(* Logix 5000 project; controller R400_500_XLS vendor 1 type 14 code 216 rev 31.11; software revision 31.01; part 14 of 32 *)
(* tags used below, declared in another part *)
   Abort1 : DINT;   // Not Used
   Alarm : SINT;   // Wait 3 seconds
   AlarmAcked : BOOL;   // Alarm has been acked
   bAlrm : BOOL[64];
   bChangeFromNonHeatedToHeated : BOOL;
   Chem_Pump : UDT_CHEM_PUMP[4];   // Chemical Pump flow rate
   CURRENT_CYCLE : DINT;
   CycExcBuffer : UDT_CYCLE;
   CycleModifBuffer : UDT_CYCLE;
   Cycles : UDT_CYCLE[11];
   DESCALER : SINT;
   ENVIRO_CARE : SINT;
   EXTRA_CARE : SINT;
   FC83_AutoSpeed : BOOL;   // Cycle pump speed selection
   FC83_AutoWtrLevel : BOOL;   // Cycle water level selection
   FC83_CyclePerm : BOOL;   // Cycle permission selection
   FC83_ONS : SINT;
   Inj_Cond : SINT;   // Conductivity injection based steps
   Inj_Time : SINT;   // Time based chemical injection steps
   M : DINT[5];   // Memory Bits
   Neutral : SINT;
   NeutralizantPump : SINT;
   NeutralizationInjTime : DINT;
   NeutralizationPhaseRequired : BOOL;
   NeutralizationRecircTime : DINT;
   ONS_WSH35 : SINT;
   PLASTIC_CARE : SINT;
   PreWash_Select : BOOL;
   PrewashIndex : SINT;   // Index of the selected pre-wash treatment
   RINSE_CARE : SINT;
   RinseIndex : SINT;
   Run : DINT;
   STANDARD : SINT;
   String : STRING[50];   // String
   Supervisor : DINT;
   Tmr : TIMER[107];
   Trt_Wsh : DINT;
   USER_DEFINED_10 : SINT;
   USER_DEFINED_11 : SINT;
   USER_DEFINED_7 : SINT;
   USER_DEFINED_8 : SINT;
   USER_DEFINED_9 : SINT;
   VolumeInjected_ML : REAL;
   VolumeNeutralizer : REAL;
   WashIndex : SINT;
   WshExcBuffer : UDT_WASH;
   cfgPrewashWport : SINT;
   CycleName : STRING[12];
   CyclePtr : DINT;   // Cycle Pointeur
   I_Chm_1_Lvl_Sw : BOOL;   // Chemical Pump #1 level switch
   I_Chm_2_Lvl_Sw : BOOL;   // Chemical Pump #2 level switch
   I_Chm_3_Lvl_Sw : BOOL;   // Chemical Pump #3 level switch
   I_Chm_4_Lvl_Sw : BOOL;   // Chemical Pump #4 level switch
   NumInputReal : UDT_NUMERIC_INPUT_REAL[17];
   Screen_Ctrl : DINT;   // PLC Screen Request
   SelChemNeutralizer : UDT_SELECTOR[5];
   Selector : UDT_SELECTOR[25];   // Piloted list selector
   Tpb : DINT[11];
   TpbImage : DINT[11];
   Unit : Hrdwre;   // Unit Configuration
(* MainProgram, continued *)

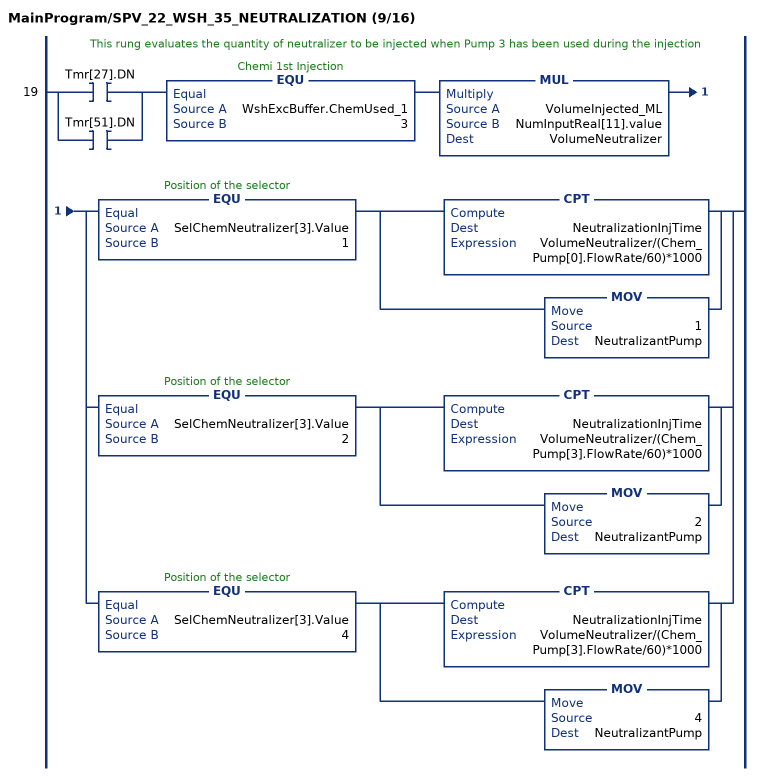
   [picture p243: MainProgram/SPV_22_WSH_35_NEUTRALIZATION rungs 19-19]
   // This rung evaluates the quantity of neutralizer to be injected when Pump 3 has been used during the injection
   19: [XIC(Tmr[27].DN) ,XIC(Tmr[51].DN) ]EQU(WshExcBuffer.ChemUsed_1,3)MUL(VolumeInjected_ML,NumInputReal[11].value,VolumeNeutralizer)[EQU(SelChemNeutralizer[3].Value,1) [CPT(NeutralizationInjTime,VolumeNeutralizer/(Chem_Pump[0].FlowRate/60)*1000) ,MOV(1,NeutralizantPump) ] ,EQU(SelChemNeutralizer[3].Value,2) [CPT(NeutralizationInjTime,VolumeNeutralizer/(Chem_Pump[3].FlowRate/60)*1000) ,MOV(2,NeutralizantPump) ] ,EQU(SelChemNeutralizer[3].Value,4) [CPT(NeutralizationInjTime,VolumeNeutralizer/(Chem_Pump[3].FlowRate/60)*1000) ,MOV(4,NeutralizantPump) ] ];
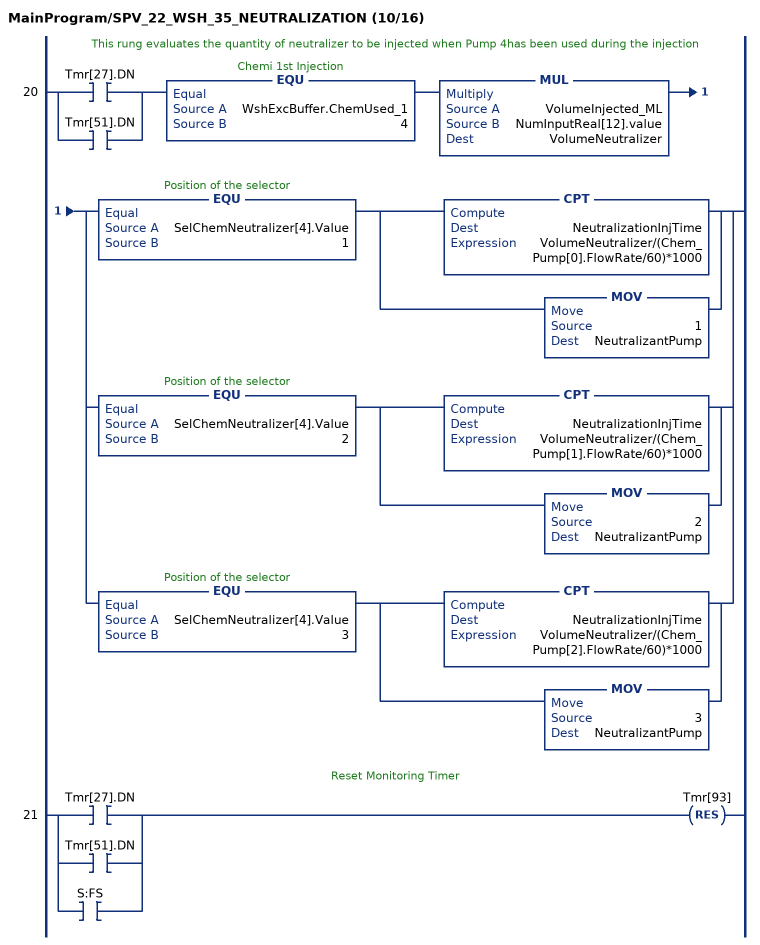
   // This rung evaluates the quantity of neutralizer to be injected when Pump 4has been used during the injection
   20: [XIC(Tmr[27].DN) ,XIC(Tmr[51].DN) ]EQU(WshExcBuffer.ChemUsed_1,4)MUL(VolumeInjected_ML,NumInputReal[12].value,VolumeNeutralizer)[EQU(SelChemNeutralizer[4].Value,1) [CPT(NeutralizationInjTime,VolumeNeutralizer/(Chem_Pump[0].FlowRate/60)*1000) ,MOV(1,NeutralizantPump) ] ,EQU(SelChemNeutralizer[4].Value,2) [CPT(NeutralizationInjTime,VolumeNeutralizer/(Chem_Pump[1].FlowRate/60)*1000) ,MOV(2,NeutralizantPump) ] ,EQU(SelChemNeutralizer[4].Value,3) [CPT(NeutralizationInjTime,VolumeNeutralizer/(Chem_Pump[2].FlowRate/60)*1000) ,MOV(3,NeutralizantPump) ] ];
   // Reset Monitoring Timer
   21: [XIC(Tmr[27].DN) ,XIC(Tmr[51].DN) ,XIC(S:FS) ]RES(Tmr[93]);
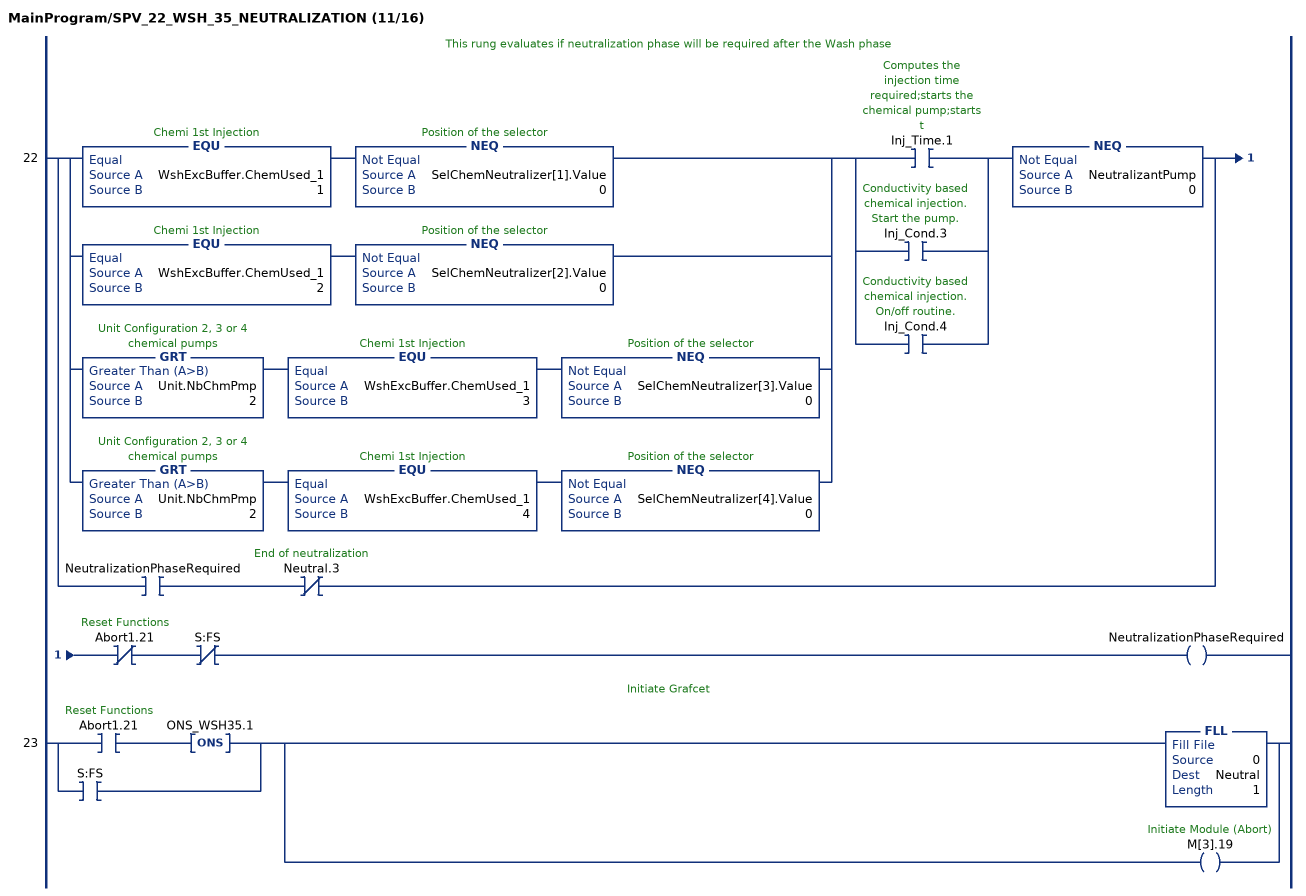
   // This rung evaluates if neutralization phase will be required after the Wash phase
   22: [[EQU(WshExcBuffer.ChemUsed_1,1) NEQ(SelChemNeutralizer[1].Value,0) ,EQU(WshExcBuffer.ChemUsed_1,2) NEQ(SelChemNeutralizer[2].Value,0) ,GRT(Unit.NbChmPmp,2) EQU(WshExcBuffer.ChemUsed_1,3) NEQ(SelChemNeutralizer[3].Value,0) ,GRT(Unit.NbChmPmp,2) EQU(WshExcBuffer.ChemUsed_1,4) NEQ(SelChemNeutralizer[4].Value,0) ] [XIC(Inj_Time.1) ,[XIC(Inj_Cond.3) ,XIC(Inj_Cond.4) ] ] NEQ(NeutralizantPump,0) ,XIC(NeutralizationPhaseRequired) XIO(Neutral.3) ]XIO(Abort1.21)XIO(S:FS)OTE(NeutralizationPhaseRequired);
   // Initiate Grafcet
   23: [XIC(Abort1.21) ONS(ONS_WSH35.1) ,XIC(S:FS) ][FLL(0,Neutral,1) ,OTE(M[3].19) ];
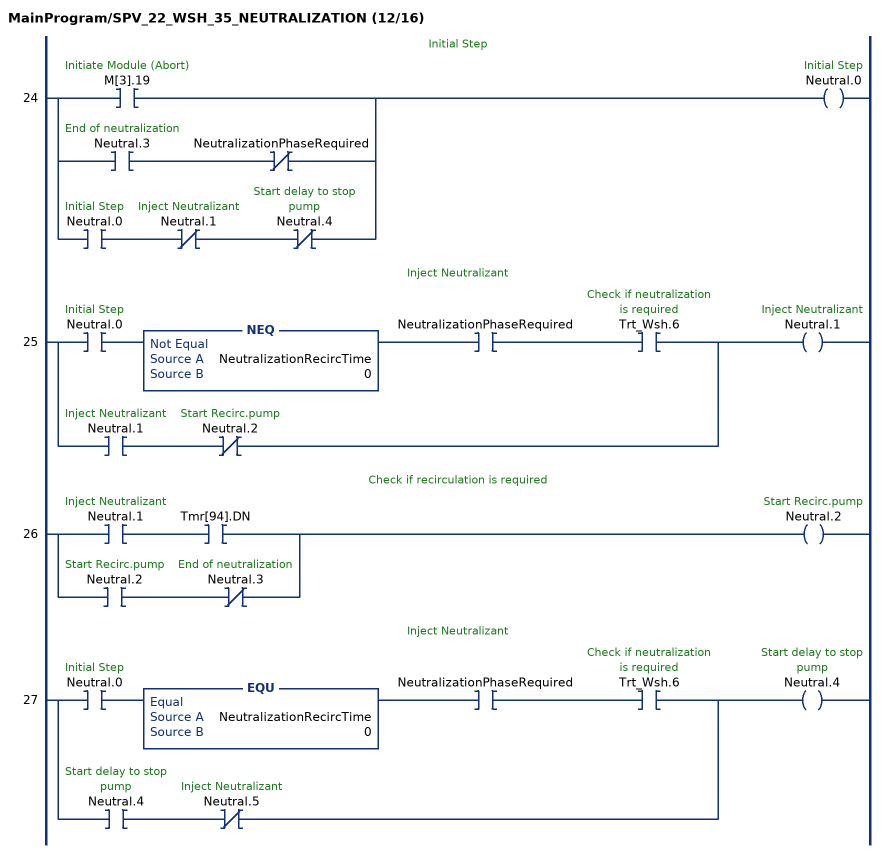
   // Initial Step
   24: [XIC(M[3].19) ,XIC(Neutral.3) XIO(NeutralizationPhaseRequired) ,XIC(Neutral.0) XIO(Neutral.1) XIO(Neutral.4) ]OTE(Neutral.0);
   // Inject Neutralizant
   25: [XIC(Neutral.0) NEQ(NeutralizationRecircTime,0) XIC(NeutralizationPhaseRequired) XIC(Trt_Wsh.6) ,XIC(Neutral.1) XIO(Neutral.2) ]OTE(Neutral.1);
   // Check if recirculation is required
   26: [XIC(Neutral.1) XIC(Tmr[94].DN) ,XIC(Neutral.2) XIO(Neutral.3) ]OTE(Neutral.2);
   // Inject Neutralizant
   27: [XIC(Neutral.0) EQU(NeutralizationRecircTime,0) XIC(NeutralizationPhaseRequired) XIC(Trt_Wsh.6) ,XIC(Neutral.4) XIO(Neutral.5) ]OTE(Neutral.4);
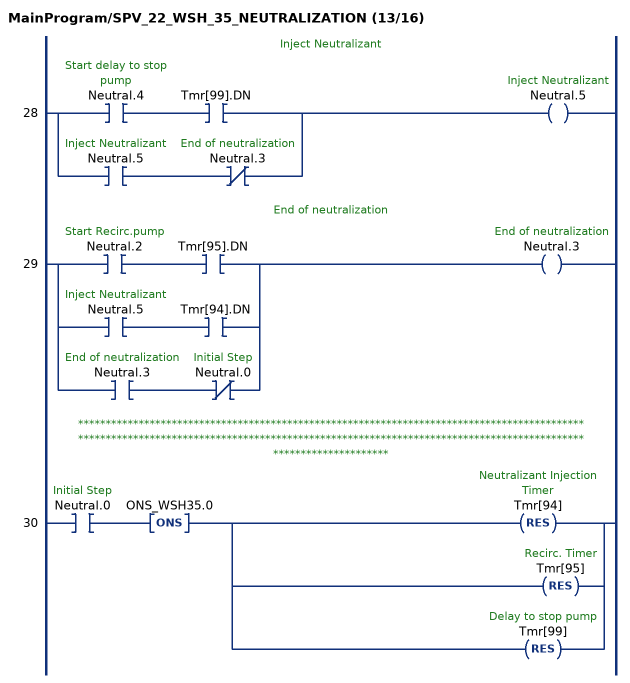
   // Inject Neutralizant
   28: [XIC(Neutral.4) XIC(Tmr[99].DN) ,XIC(Neutral.5) XIO(Neutral.3) ]OTE(Neutral.5);
   // End of neutralization
   29: [XIC(Neutral.2) XIC(Tmr[95].DN) ,XIC(Neutral.5) XIC(Tmr[94].DN) ,XIC(Neutral.3) XIO(Neutral.0) ]OTE(Neutral.3);
   // *************************************************************************************************************************************************************************************************************
   30: XIC(Neutral.0)ONS(ONS_WSH35.0)[RES(Tmr[94]) ,RES(Tmr[95]) ,RES(Tmr[99]) ];
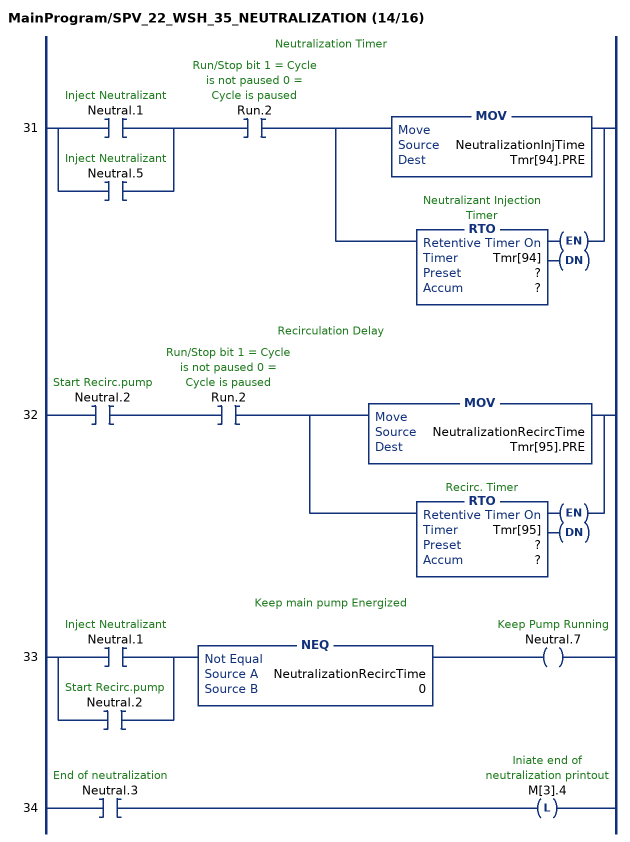
   // Neutralization Timer
   31: [XIC(Neutral.1) ,XIC(Neutral.5) ]XIC(Run.2)[MOV(NeutralizationInjTime,Tmr[94].PRE) ,RTO(Tmr[94],?,?) ];
   // Recirculation Delay
   32: XIC(Neutral.2)XIC(Run.2)[MOV(NeutralizationRecircTime,Tmr[95].PRE) ,RTO(Tmr[95],?,?) ];
   // Keep main pump Energized
   33: [XIC(Neutral.1) ,XIC(Neutral.2) ]NEQ(NeutralizationRecircTime,0)OTE(Neutral.7);
   34: XIC(Neutral.3)OTL(M[3].4);
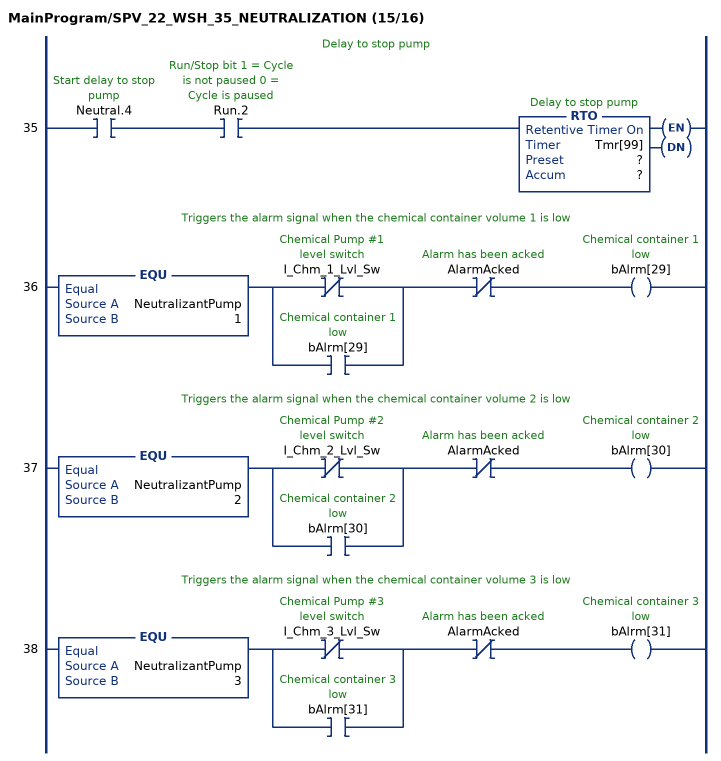
   // Delay to stop pump
   35: XIC(Neutral.4)XIC(Run.2)RTO(Tmr[99],?,?);
   // Triggers the alarm signal when the chemical container volume 1 is low
   36: EQU(NeutralizantPump,1)[XIO(I_Chm_1_Lvl_Sw) ,XIC(bAlrm[29]) ]XIO(AlarmAcked)OTE(bAlrm[29]);
   // Triggers the alarm signal when the chemical container volume 2 is low
   37: EQU(NeutralizantPump,2)[XIO(I_Chm_2_Lvl_Sw) ,XIC(bAlrm[30]) ]XIO(AlarmAcked)OTE(bAlrm[30]);
   // Triggers the alarm signal when the chemical container volume 3 is low
   38: EQU(NeutralizantPump,3)[XIO(I_Chm_3_Lvl_Sw) ,XIC(bAlrm[31]) ]XIO(AlarmAcked)OTE(bAlrm[31]);
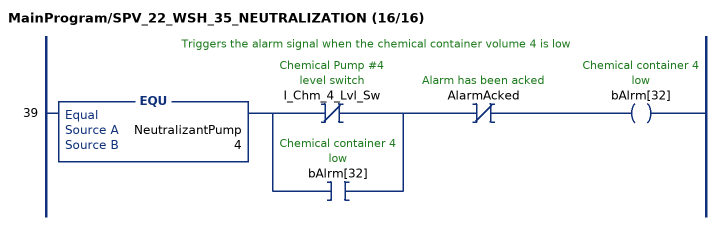
   // Triggers the alarm signal when the chemical container volume 4 is low
   39: EQU(NeutralizantPump,4)[XIO(I_Chm_4_Lvl_Sw) ,XIC(bAlrm[32]) ]XIO(AlarmAcked)OTE(bAlrm[32]);
END_ROUTINE

ROUTINE SPV_3_5_6_7_13_14_15_CYC_MOD   (* ladder *)
// This routine manages the HMI screens and the logic in order for the supervisor to modify the cycle parameters
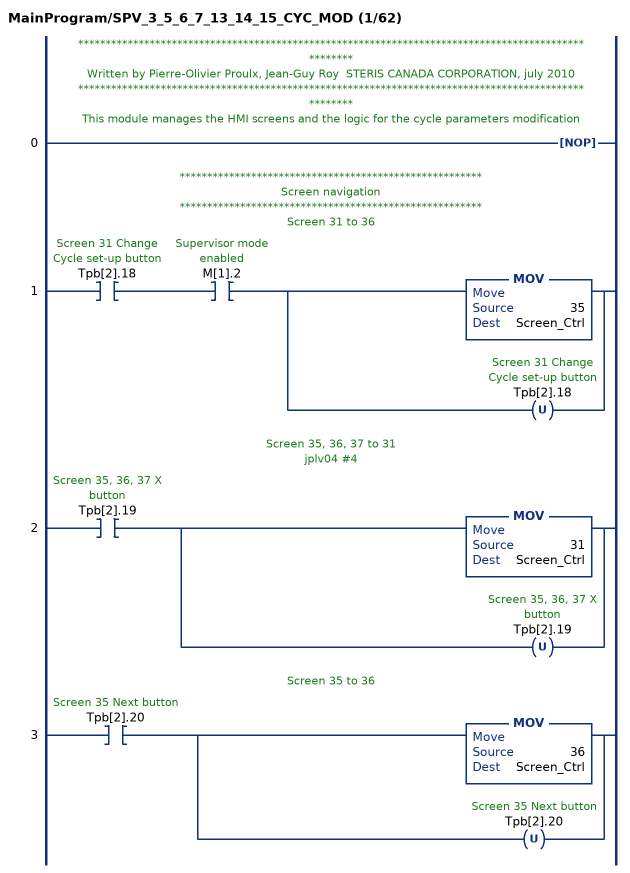
   // ****************************************************************************************************
   // Written by Pierre-Olivier Proulx, Jean-Guy Roy  STERIS CANADA CORPORATION, july 2010
   // ****************************************************************************************************
   // This module manages the HMI screens and the logic for the cycle parameters modification
   0: NOP();
   // *******************************************************
   // Screen navigation
   // *******************************************************
   // Screen 31 to 36
   1: XIC(Tpb[2].18)XIC(M[1].2)[MOV(35,Screen_Ctrl) ,OTU(Tpb[2].18) ];
   // Screen 35, 36, 37 to 31
   // jplv04 #4
   2: XIC(Tpb[2].19)[MOV(31,Screen_Ctrl) ,OTU(Tpb[2].19) ];
   // Screen 35 to 36
   3: XIC(Tpb[2].20)[MOV(36,Screen_Ctrl) ,OTU(Tpb[2].20) ];
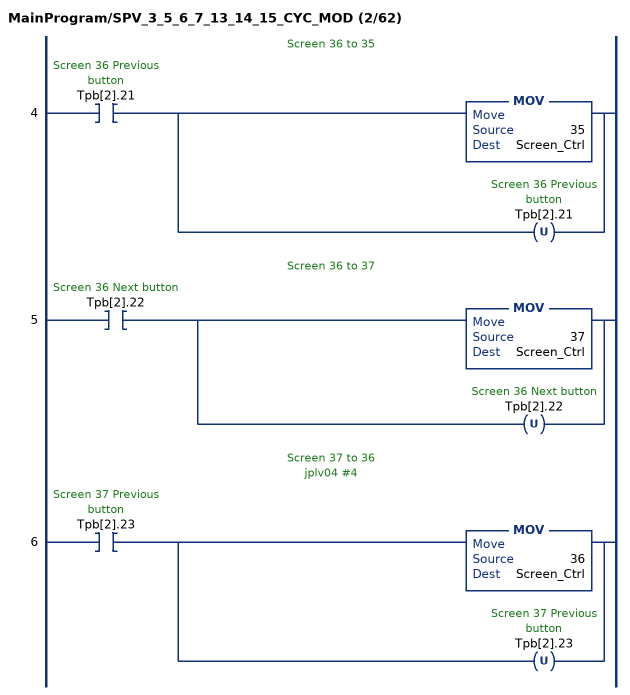
   // Screen 36 to 35
   4: XIC(Tpb[2].21)[MOV(35,Screen_Ctrl) ,OTU(Tpb[2].21) ];
   // Screen 36 to 37
   5: XIC(Tpb[2].22)[MOV(37,Screen_Ctrl) ,OTU(Tpb[2].22) ];
   // Screen 37 to 36
   // jplv04 #4
   6: XIC(Tpb[2].23)[MOV(36,Screen_Ctrl) ,OTU(Tpb[2].23) ];
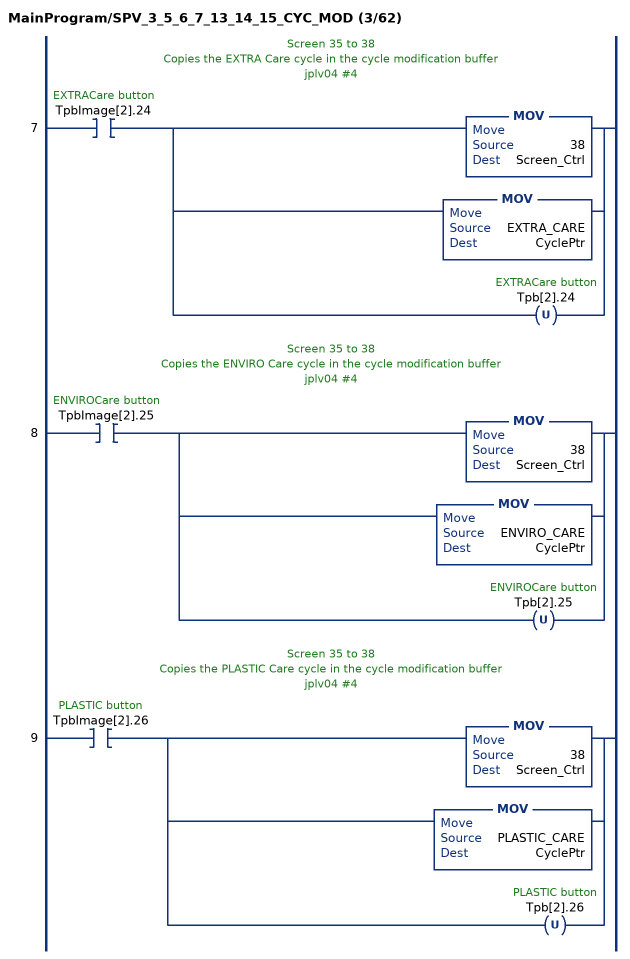
   // Screen 35 to 38
   // Copies the EXTRA Care cycle in the cycle modification buffer
   // jplv04 #4
   7: XIC(TpbImage[2].24)[MOV(38,Screen_Ctrl) ,MOV(EXTRA_CARE,CyclePtr) ,OTU(Tpb[2].24) ];
   // Screen 35 to 38
   // Copies the ENVIRO Care cycle in the cycle modification buffer
   // jplv04 #4
   8: XIC(TpbImage[2].25)[MOV(38,Screen_Ctrl) ,MOV(ENVIRO_CARE,CyclePtr) ,OTU(Tpb[2].25) ];
   // Screen 35 to 38
   // Copies the PLASTIC Care cycle in the cycle modification buffer
   // jplv04 #4
   9: XIC(TpbImage[2].26)[MOV(38,Screen_Ctrl) ,MOV(PLASTIC_CARE,CyclePtr) ,OTU(Tpb[2].26) ];
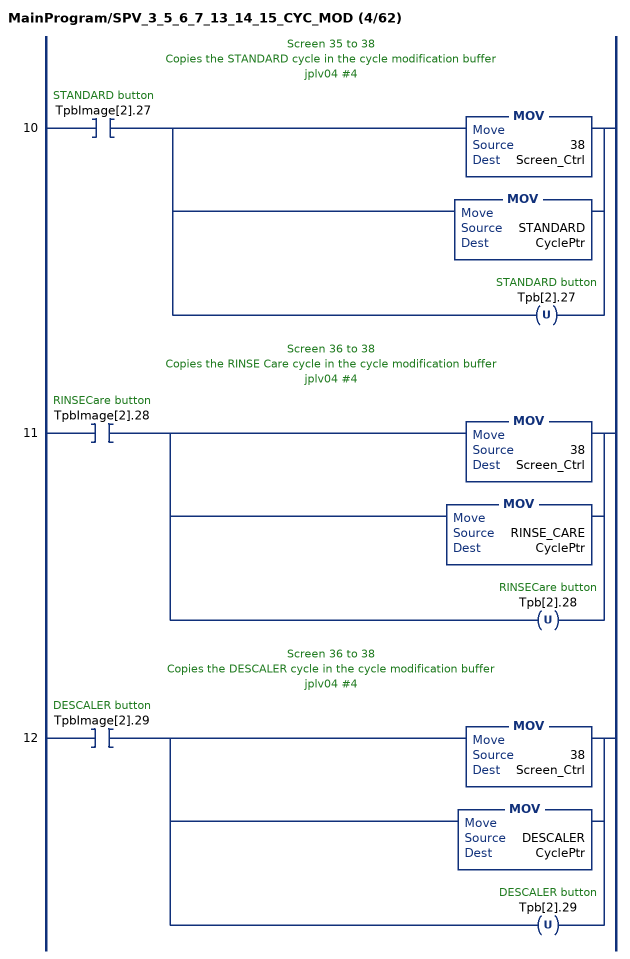
   // Screen 35 to 38
   // Copies the STANDARD cycle in the cycle modification buffer
   // jplv04 #4
   10: XIC(TpbImage[2].27)[MOV(38,Screen_Ctrl) ,MOV(STANDARD,CyclePtr) ,OTU(Tpb[2].27) ];
   // Screen 36 to 38
   // Copies the RINSE Care cycle in the cycle modification buffer
   // jplv04 #4
   11: XIC(TpbImage[2].28)[MOV(38,Screen_Ctrl) ,MOV(RINSE_CARE,CyclePtr) ,OTU(Tpb[2].28) ];
   // Screen 36 to 38
   // Copies the DESCALER cycle in the cycle modification buffer
   // jplv04 #4
   12: XIC(TpbImage[2].29)[MOV(38,Screen_Ctrl) ,MOV(DESCALER,CyclePtr) ,OTU(Tpb[2].29) ];
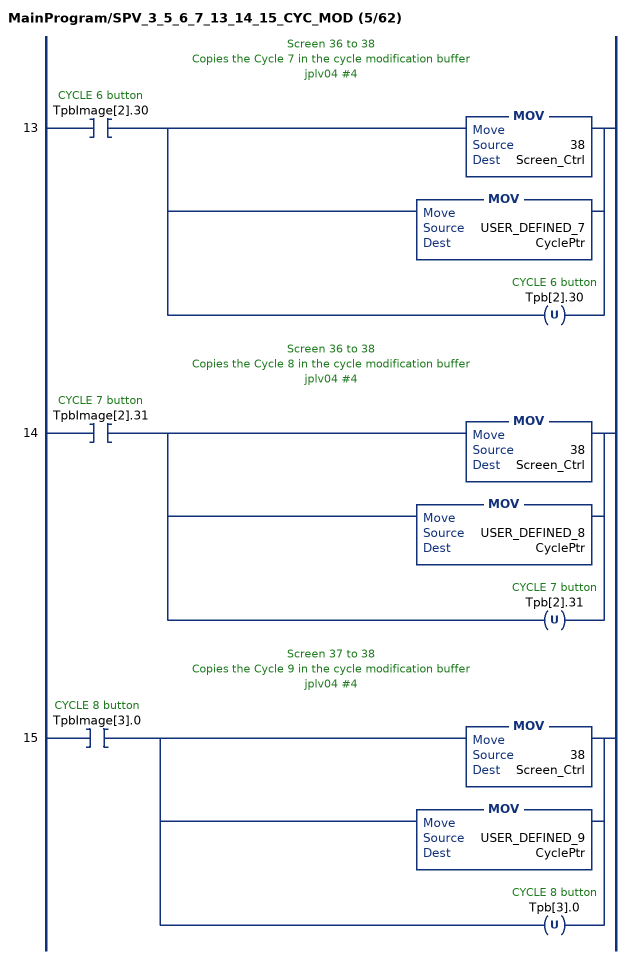
   // Screen 36 to 38
   // Copies the Cycle 7 in the cycle modification buffer
   // jplv04 #4
   13: XIC(TpbImage[2].30)[MOV(38,Screen_Ctrl) ,MOV(USER_DEFINED_7,CyclePtr) ,OTU(Tpb[2].30) ];
   // Screen 36 to 38
   // Copies the Cycle 8 in the cycle modification buffer
   // jplv04 #4
   14: XIC(TpbImage[2].31)[MOV(38,Screen_Ctrl) ,MOV(USER_DEFINED_8,CyclePtr) ,OTU(Tpb[2].31) ];
   // Screen 37 to 38
   // Copies the Cycle 9 in the cycle modification buffer
   // jplv04 #4
   15: XIC(TpbImage[3].0)[MOV(38,Screen_Ctrl) ,MOV(USER_DEFINED_9,CyclePtr) ,OTU(Tpb[3].0) ];
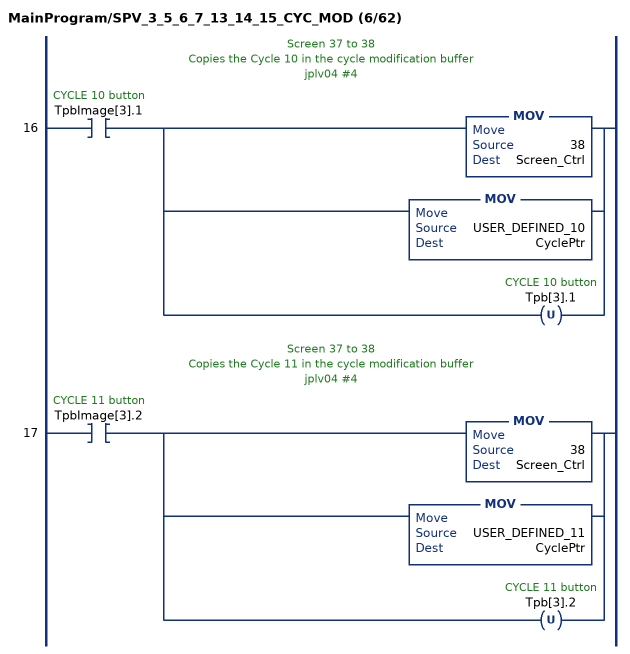
   // Screen 37 to 38
   // Copies the Cycle 10 in the cycle modification buffer
   // jplv04 #4
   16: XIC(TpbImage[3].1)[MOV(38,Screen_Ctrl) ,MOV(USER_DEFINED_10,CyclePtr) ,OTU(Tpb[3].1) ];
   // Screen 37 to 38
   // Copies the Cycle 11 in the cycle modification buffer
   // jplv04 #4
   17: XIC(TpbImage[3].2)[MOV(38,Screen_Ctrl) ,MOV(USER_DEFINED_11,CyclePtr) ,OTU(Tpb[3].2) ];
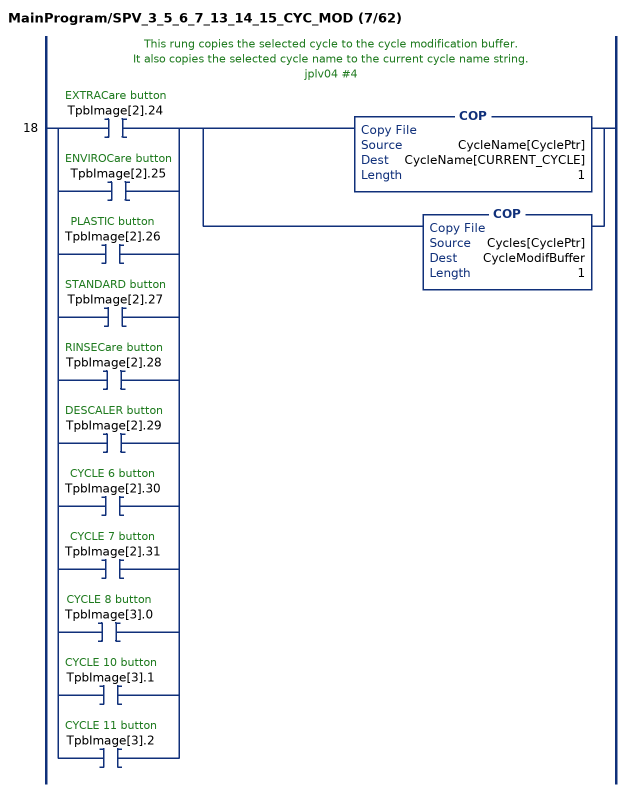
   // This rung copies the selected cycle to the cycle modification buffer.
   // It also copies the selected cycle name to the current cycle name string.
   // jplv04 #4
   18: [XIC(TpbImage[2].24) ,XIC(TpbImage[2].25) ,XIC(TpbImage[2].26) ,XIC(TpbImage[2].27) ,XIC(TpbImage[2].28) ,XIC(TpbImage[2].29) ,XIC(TpbImage[2].30) ,XIC(TpbImage[2].31) ,XIC(TpbImage[3].0) ,XIC(TpbImage[3].1) ,XIC(TpbImage[3].2) ][COP(CycleName[CyclePtr],CycleName[CURRENT_CYCLE],1) ,COP(Cycles[CyclePtr],CycleModifBuffer,1) ];
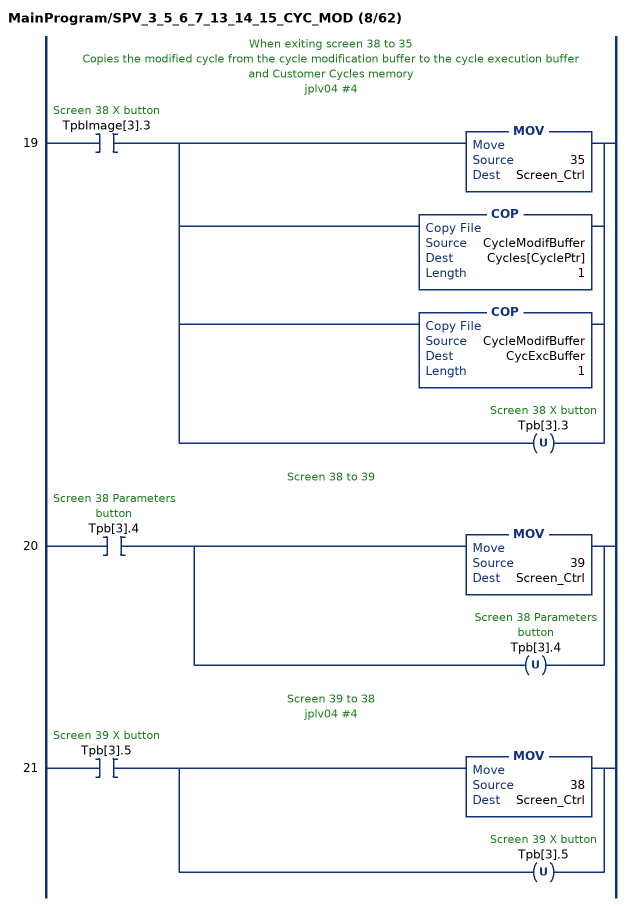
   // When exiting screen 38 to 35
   // Copies the modified cycle from the cycle modification buffer to the cycle execution buffer and Customer Cycles memory
   // jplv04 #4
   19: XIC(TpbImage[3].3)[MOV(35,Screen_Ctrl) ,COP(CycleModifBuffer,Cycles[CyclePtr],1) ,COP(CycleModifBuffer,CycExcBuffer,1) ,OTU(Tpb[3].3) ];
   // Screen 38 to 39
   20: XIC(Tpb[3].4)[MOV(39,Screen_Ctrl) ,OTU(Tpb[3].4) ];
   // Screen 39 to 38
   // jplv04 #4
   21: XIC(Tpb[3].5)[MOV(38,Screen_Ctrl) ,OTU(Tpb[3].5) ];
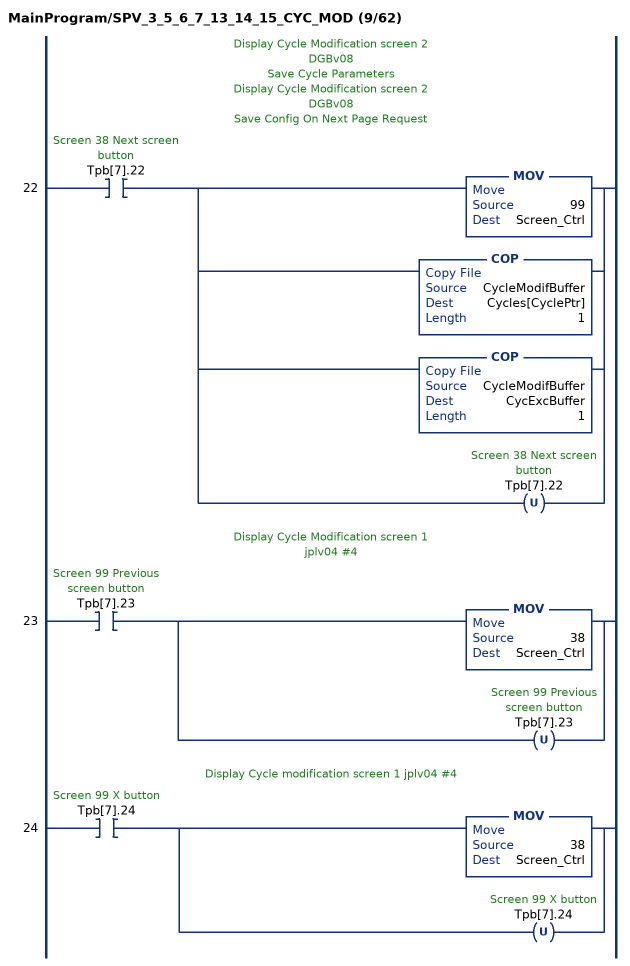
   // Display Cycle Modification screen 2
   // DGBv08
   // Save Cycle Parameters
   // Display Cycle Modification screen 2
   // DGBv08
   // Save Config On Next Page Request
   22: XIC(Tpb[7].22)[MOV(99,Screen_Ctrl) ,COP(CycleModifBuffer,Cycles[CyclePtr],1) ,COP(CycleModifBuffer,CycExcBuffer,1) ,OTU(Tpb[7].22) ];
   // Display Cycle Modification screen 1
   // jplv04 #4
   23: XIC(Tpb[7].23)[MOV(38,Screen_Ctrl) ,OTU(Tpb[7].23) ];
   // Display Cycle modification screen 1 jplv04 #4
   24: XIC(Tpb[7].24)[MOV(38,Screen_Ctrl) ,OTU(Tpb[7].24) ];
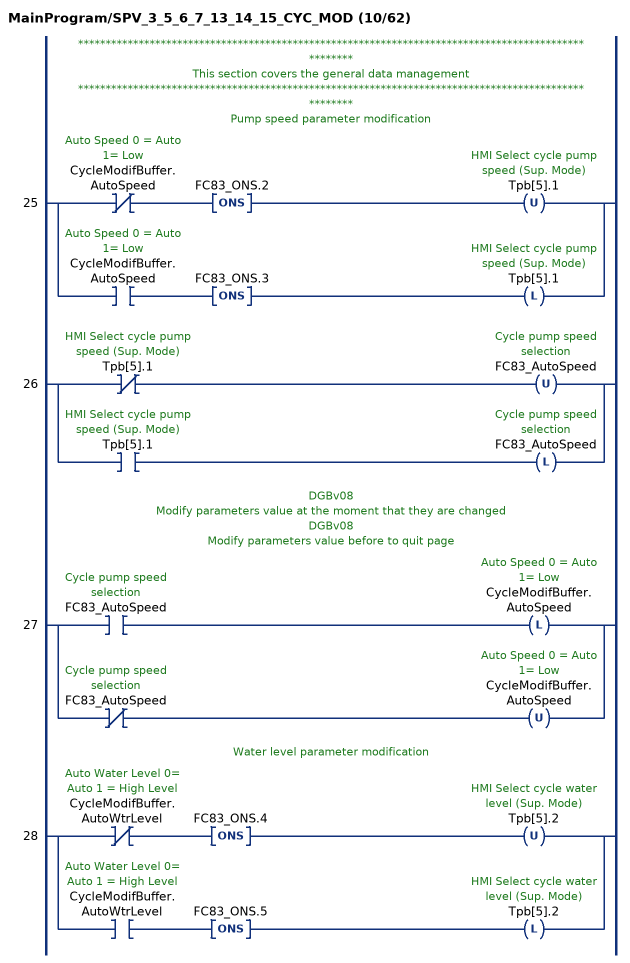
   // ****************************************************************************************************
   // This section covers the general data management
   // ****************************************************************************************************
   // Pump speed parameter modification
   25: [XIO(CycleModifBuffer.AutoSpeed) ONS(FC83_ONS.2) OTU(Tpb[5].1) ,XIC(CycleModifBuffer.AutoSpeed) ONS(FC83_ONS.3) OTL(Tpb[5].1) ];
   26: [XIO(Tpb[5].1) OTU(FC83_AutoSpeed) ,XIC(Tpb[5].1) OTL(FC83_AutoSpeed) ];
   // DGBv08
   // Modify parameters value at the moment that they are changed
   // DGBv08
   // Modify parameters value before to quit page
   27: [XIC(FC83_AutoSpeed) OTL(CycleModifBuffer.AutoSpeed) ,XIO(FC83_AutoSpeed) OTU(CycleModifBuffer.AutoSpeed) ];
   // Water level parameter modification
   28: [XIO(CycleModifBuffer.AutoWtrLevel) ONS(FC83_ONS.4) OTU(Tpb[5].2) ,XIC(CycleModifBuffer.AutoWtrLevel) ONS(FC83_ONS.5) OTL(Tpb[5].2) ];
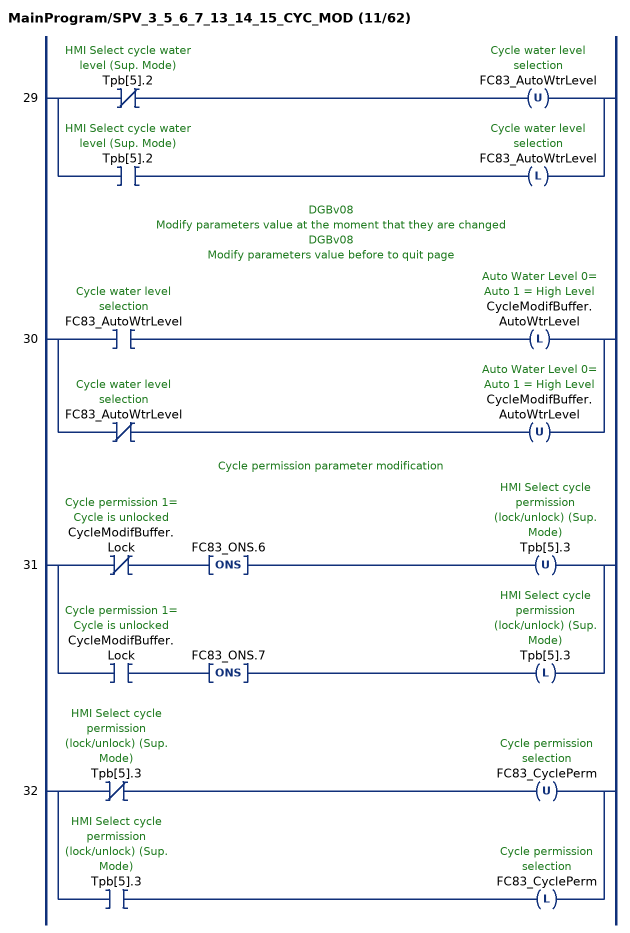
   29: [XIO(Tpb[5].2) OTU(FC83_AutoWtrLevel) ,XIC(Tpb[5].2) OTL(FC83_AutoWtrLevel) ];
   // DGBv08
   // Modify parameters value at the moment that they are changed
   // DGBv08
   // Modify parameters value before to quit page
   30: [XIC(FC83_AutoWtrLevel) OTL(CycleModifBuffer.AutoWtrLevel) ,XIO(FC83_AutoWtrLevel) OTU(CycleModifBuffer.AutoWtrLevel) ];
   // Cycle permission parameter modification
   31: [XIO(CycleModifBuffer.Lock) ONS(FC83_ONS.6) OTU(Tpb[5].3) ,XIC(CycleModifBuffer.Lock) ONS(FC83_ONS.7) OTL(Tpb[5].3) ];
   32: [XIO(Tpb[5].3) OTU(FC83_CyclePerm) ,XIC(Tpb[5].3) OTL(FC83_CyclePerm) ];
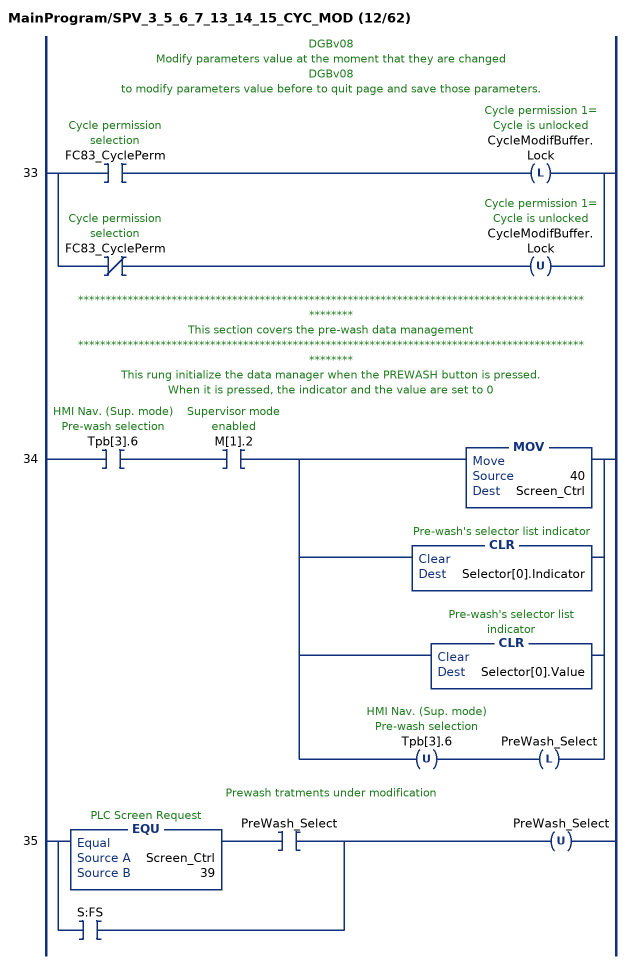
   // DGBv08
   // Modify parameters value at the moment that they are changed
   // DGBv08
   // to modify parameters value before to quit page and save those parameters.
   33: [XIC(FC83_CyclePerm) OTL(CycleModifBuffer.Lock) ,XIO(FC83_CyclePerm) OTU(CycleModifBuffer.Lock) ];
   // ****************************************************************************************************
   // This section covers the pre-wash data management
   // ****************************************************************************************************
   // This rung initialize the data manager when the PREWASH button is pressed.
   // When it is pressed, the indicator and the value are set to 0
   34: XIC(Tpb[3].6)XIC(M[1].2)[MOV(40,Screen_Ctrl) ,CLR(Selector[0].Indicator) ,CLR(Selector[0].Value) ,OTU(Tpb[3].6) OTL(PreWash_Select) ];
   // Prewash tratments under modification
   35: [EQU(Screen_Ctrl,39) XIC(PreWash_Select) ,XIC(S:FS) ]OTU(PreWash_Select);
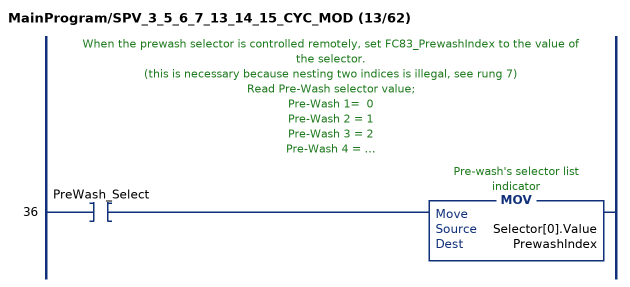
   // When the prewash selector is controlled remotely, set FC83_PrewashIndex to the value of the selector.
   // (this is necessary because nesting two indices is illegal, see rung 7)
   // Read Pre-Wash selector value;
   // Pre-Wash 1=  0
   // Pre-Wash 2 = 1
   // Pre-Wash 3 = 2
   // Pre-Wash 4 = 3
   // XLSV10  DGB  2018-09-04 : Aded Wash 3 & 4
   36: XIC(PreWash_Select)MOV(Selector[0].Value,PrewashIndex);
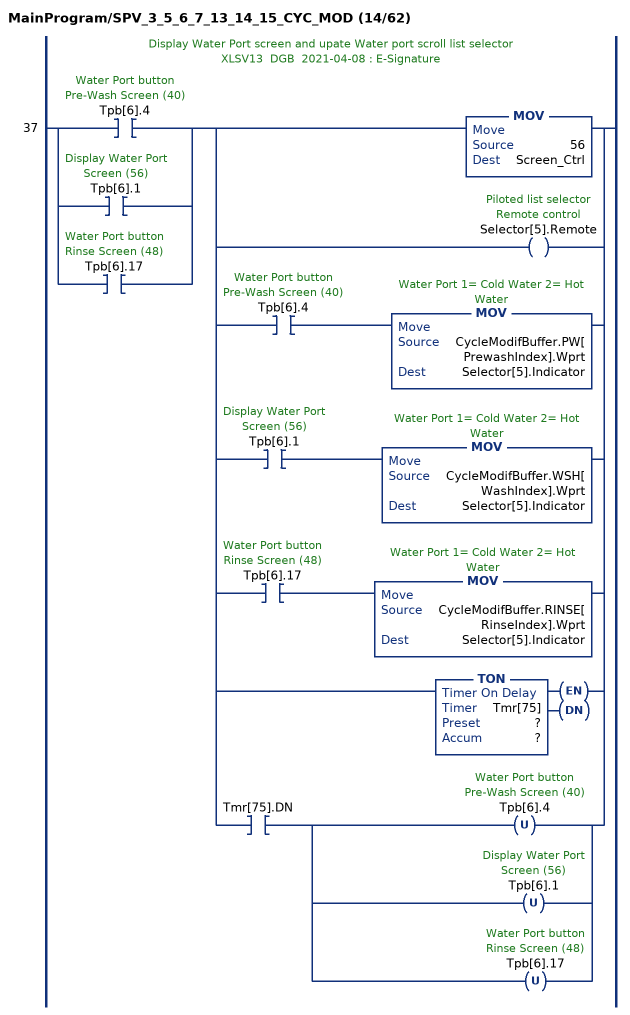
   // Display Water Port screen and upate Water port scroll list selector
   // XLSV13  DGB  2021-04-08 : E-Signature
   37: [XIC(Tpb[6].4) ,XIC(Tpb[6].1) ,XIC(Tpb[6].17) ][MOV(56,Screen_Ctrl) ,OTE(Selector[5].Remote) ,XIC(Tpb[6].4) MOV(CycleModifBuffer.PW[PrewashIndex].Wprt,Selector[5].Indicator) ,XIC(Tpb[6].1) MOV(CycleModifBuffer.WSH[WashIndex].Wprt,Selector[5].Indicator) ,XIC(Tpb[6].17) MOV(CycleModifBuffer.RINSE[RinseIndex].Wprt,Selector[5].Indicator) ,TON(Tmr[75],?,?) ,XIC(Tmr[75].DN) [OTU(Tpb[6].4) ,OTU(Tpb[6].1) ,OTU(Tpb[6].17) ] ];
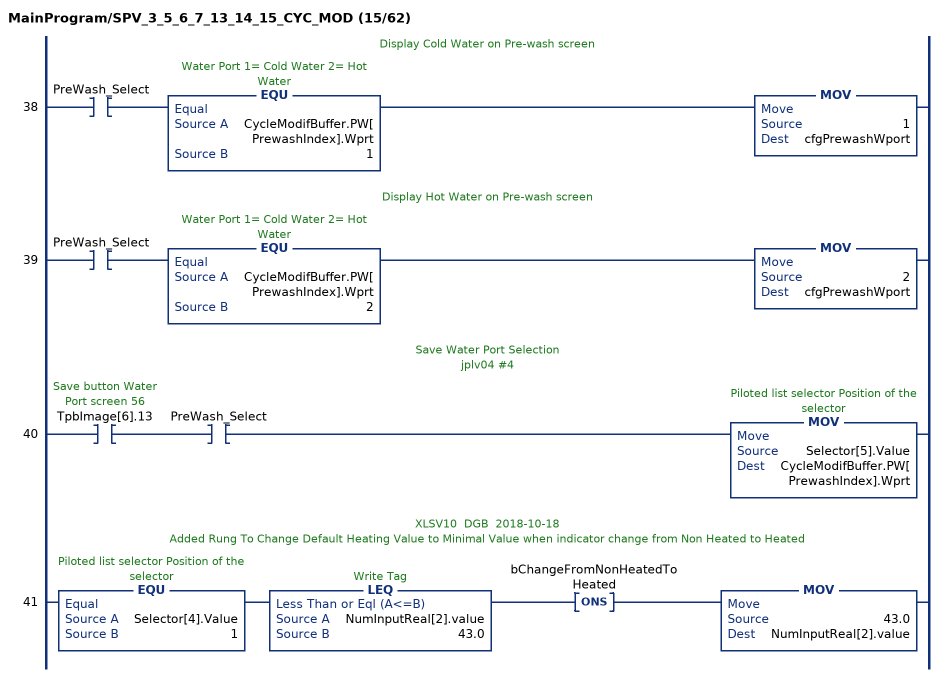
   // Display Cold Water on Pre-wash screen
   38: XIC(PreWash_Select)EQU(CycleModifBuffer.PW[PrewashIndex].Wprt,1)MOV(1,cfgPrewashWport);
   // Display Hot Water on Pre-wash screen
   39: XIC(PreWash_Select)EQU(CycleModifBuffer.PW[PrewashIndex].Wprt,2)MOV(2,cfgPrewashWport);
   // Save Water Port Selection
   // jplv04 #4
   40: XIC(TpbImage[6].13)XIC(PreWash_Select)MOV(Selector[5].Value,CycleModifBuffer.PW[PrewashIndex].Wprt);
   // XLSV10  DGB  2018-10-18
   // Added Rung To Change Default Heating Value to Minimal Value when indicator change from Non Heated to Heated
   41: EQU(Selector[4].Value,1)LEQ(NumInputReal[2].value,43.0)ONS(bChangeFromNonHeatedToHeated)MOV(43.0,NumInputReal[2].value);
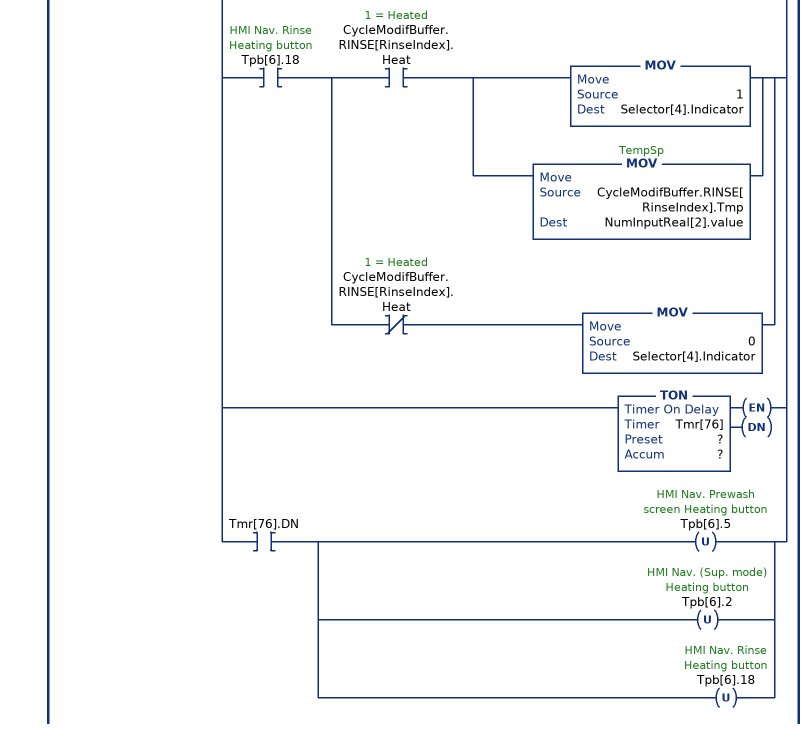
   // Prewash configuration, Display Heating screen
   // XLSV13  DGB  2021-04-08 : E-Signature
   42: [XIC(Tpb[6].5) ,XIC(Tpb[6].2) ,XIC(Tpb[6].18) ][MOV(57,Screen_Ctrl) ,OTE(Selector[4].Remote) ,XIC(Tpb[6].5) [XIC(CycleModifBuffer.PW[PrewashIndex].Heat) [MOV(1,Selector[4].Indicator) ,MOV(CycleModifBuffer.PW[PrewashIndex].Tmp,NumInputReal[2].value) ] ,XIO(CycleModifBuffer.PW[PrewashIndex].Heat) MOV(0,Selector[4].Indicator) ] ,XIC(Tpb[6].2) [XIC(CycleModifBuffer.WSH[WashIndex].Heat) [MOV(1,Selector[4].Indicator) ,MOV(CycleModifBuffer.WSH[WashIndex].Tmp,NumInputReal[2].value) ] ,XIO(CycleModifBuffer.WSH[WashIndex].Heat) MOV(0,Selector[4].Indicator) ] ,XIC(Tpb[6].18) [XIC(CycleModifBuffer.RINSE[RinseIndex].Heat) [MOV(1,Selector[4].Indicator) ,MOV(CycleModifBuffer.RINSE[RinseIndex].Tmp,NumInputReal[2].value) ] ,XIO(CycleModifBuffer.RINSE[RinseIndex].Heat) MOV(0,Selector[4].Indicator) ] ,TON(Tmr[76],?,?) ,XIC(Tmr[76].DN) [OTU(Tpb[6].5) ,OTU(Tpb[6].2) ,OTU(Tpb[6].18) ] ];
